// TIA Portal V20 export
// export: Created 2026-10-20T12:40:00.8102062Z, ExportSetting WithDefaults, DisplayName Totally Integrated Automation Portal, DisplayVersion V20 Update 6, DisplayName TIA Portal Openness, DisplayVersion V20 Update 6, DisplayName TIA Portal Version Control Interface, DisplayVersion V20 Update 6, DisplayName SINAMICS Startdrive Advanced, DisplayVersion V20 SP1, DisplayName SINAMICS Startdrive G130, G150, S120, S150, SINAMICS MV, G220, S200, S210, DisplayVersion V20 SP1, DisplayName SINAMICS Startdrive G110M, G120, G120C, G120D, G120P, G115D, DisplayVersion V20 SP1, DisplayName STEP 7 Professional, DisplayVersion V20 Update 6, DisplayName STEP 7 Safety, DisplayVersion V20 Update 2, DisplayName WinCC Basic/Comfort/Advanced, DisplayVersion V20 Update 6, DisplayName WinCC Unified, DisplayVersion V20 Update 6
DATA_BLOCK "VTD_FB_DB_4"   // DB165
VERSION : 0.1
// stored: AutoNumber true, DBAccessibleFromOPCUA true, InstanceOfName VTD_FB, InstanceOfType FB
"VTD_FB"
   // VAR_INPUT
   //    System_no : UInt;
   //    Safety_OK_Delayed : Bool;
   //    Safety_OK : Bool;
   //    Cnv_Sensors : "Cnv_Inputs";
   //    VTD_Settings : "VTD_Settings";
   //    Bypass_LP : Bool;
   //    Bypass : "Safety_Bypass_RemotePanel";
   // END_VAR
   // VAR_IN_OUT
   //    VTD_Control : "VTD_Control";
   //    SinaSpeed : SinaSpeed;
   //    LE_Bypass_HMI : Bool;
   // END_VAR
   // VAR
   //    State : UInt;
   //    Last_State : UInt;
   //    I_State : UInt;
   //    LD_Timer_1 : TON_TIME;
   //    LD_Timer : TON_TIME;
   //    DP_Timer { S7_SetPoint := 'True'} : TON_TIME;
   //    Watchdog { S7_SetPoint := 'True'} : TON_TIME;
   //    CS_TImer { S7_SetPoint := 'True'} : TON_TIME;
   //    Interlock_Timer { S7_SetPoint := 'True'} : TON_TIME;
   //    MainSetpoint : Int;
   //    Position_Offset : Real;
   //    ChangeToLow : Array[1..4] of DInt;
   //    DestPosition : Real;
   //    SetUpSpeed : UInt;
   //    LevelBelowExtractor : UInt;
   //    IEC_Timer_0_Instance { S7_SetPoint := 'True'} : TON_TIME;
   //    DestinationLevel : UInt;
   //    CurrentlLevel : UInt;
   //    VTD_ID_Decoded { ExternalAccessible := 'False'; ExternalVisible := 'False'; ExternalWritable := 'False'} : "ID_Decoded";
   //    Cnv_ID_Decoded { ExternalAccessible := 'False'; ExternalVisible := 'False'; ExternalWritable := 'False'} : Array[1..2] of "ID_Decoded";
   //    IEC_Timer_0_Instance_1 { S7_SetPoint := 'True'} : TON_TIME;
   //    IEC_Timer_0_Instance_2 { S7_SetPoint := 'True'} : TON_TIME;
   //    VTD_ControlInstructionTask_ID_Old : Int;
   //    R_Execulte { S7_SetPoint := 'True'} : R_TRIG;
   //    R_AutomatcMode { S7_SetPoint := 'True'} : R_TRIG;
   //    T_Encoders_Difference { S7_SetPoint := 'True'} : TON_TIME;
   //    T_LE_Error { S7_SetPoint := 'True'} : TON_TIME;
   //    T_Setpoint_Delay { S7_SetPoint := 'True'} : TON_TIME;
   //    Distance_mm : Real;
   //    TravelTime_s : UInt;
   //    LE_Prev_mm : Real;
   //    DeltaPos_mm : Real;
   //    SampleTime_s : Real;
   //    VTDSpeed_mm_s : Real;
   //    T_Speed { S7_SetPoint := 'True'} : TON_TIME;
   //    Speed_mm_per_percent : Real;
   //    Speed_mm_s { ExternalAccessible := 'False'; ExternalVisible := 'False'; ExternalWritable := 'False'} : Real;
   //    TravelTime_ms { ExternalAccessible := 'False'; ExternalVisible := 'False'; ExternalWritable := 'False'} : UInt;
   //    Watchdog_PT { ExternalAccessible := 'False'; ExternalVisible := 'False'; ExternalWritable := 'False'} : Time;
   //    Stopper_Extend_Timer { S7_SetPoint := 'True'} : TON_TIME;
   //    T_LE_read_0 { S7_SetPoint := 'True'} : TON_TIME;
   // END_VAR
BEGIN
END_DATA_BLOCK
